FUNCTION_BLOCK PRINT_START
  {SET_ATTRIBUTE(OpcUa, SERVICE)}
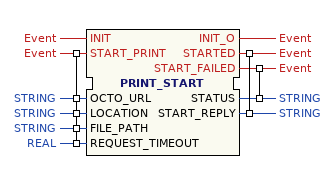
  EVENT_INPUT
    INIT;
    START_PRINT WITH OCTO_URL, LOCATION, FILE_PATH, REQUEST_TIMEOUT;
  END_EVENT
  EVENT_OUTPUT
    INIT_O;
    STARTED WITH START_REPLY;
    START_FAILED WITH STATUS;
  END_EVENT
  VAR_INPUT
    OCTO_URL : STRING; {SET_ATTRIBUTE(OpcUa, Constant)}
    LOCATION : STRING; {SET_ATTRIBUTE(OpcUa, Constant)}
    FILE_PATH : STRING; {SET_ATTRIBUTE(OpcUa, Variable)}
    REQUEST_TIMEOUT : REAL; {SET_ATTRIBUTE(OpcUa, Constant)}
  END_VAR
  VAR_OUTPUT
    STATUS : STRING; {SET_ATTRIBUTE(OpcUa, Variable)}
    START_REPLY : STRING; {SET_ATTRIBUTE(OpcUa, Variable)}
  END_VAR
END_FUNCTION_BLOCK
